Universal Robots PolyScope program: test.urp

Program test (installation=default directory=/programs createdIn=5.23.0 lastSavedIn=5.23.0 robotSerialNumber=20245590068)
Calibrated DH parameters: a=[0.00013, -0.03651, -0.389144, 0.000102, 0.000008, 0]; d=[0.162613, 192.230671, -179.915756, -12.181517, 0.099698, 0.099535]; alpha=[1.57038, 0.002205, 0.004138, 1.570804, -1.571025, 0]; deltaTheta=[-0.000001, 1.484886, 4.928506, -0.130209, 0, 0]
InitVariablesNode
Robot Program (runOnlyOnce=false)
  Popup Message (haltProgram=false message=robot moving inputType=Text)
  Loop Counting (count=5) loopVariable(name=Loop_1)
    MoveL speed 250 mm/s, acceleration 1200 mm/s^2 (useActiveTCP=true optimoveEnabled=false optiMoveSpeed=0.3 optiMoveAcceleration=0.09) feature=Base
      MoveDirectionNode (selectedDirection=ZMinus toolParams=0.05, 0.1)
        Until DISTANCE (allowActions=false deceleration=3 distanceNodeType=STOP) Distance=0.001; motionParameters(blendRadius=0)
      Wait Sleep waitTime=10
